(*
SPDX-FileCopyrightText: © 2026 Oleksandr Tiutyk <trofimich@gmail.com>
SPDX-License-Identifier: MIT
License: https://opensource.org/license/mit
*)

(*!
<summary>
Beckhoff EL1512: 2-channel up/down counter terminal (24 V DC).
</summary>
<description>
Represents the default 2Ch. Counter assignment: TxPDOs 0x1A00/0x1A01 and RxPDOs 0x1600/0x1601.
Each channel has 16-bit status/control and a 32-bit counter/preset. Direction is configured through CoE.
Single-channel up/down or gated-counter assignments are outside this model.
When used for I/O, link located fields or their containing buffers to the matching selected PDOs.
The record is not a packed wire buffer; compiler padding is not part of the device specification.
Unlinked/default values do not prove valid I/O. The caller evaluates bus/channel validity before use.
Use one owner task per instance and externally synchronize other access; multi-field snapshots are not atomic.
Copies store data without creating hardware links. Keep borrowed field references valid while consumers are bound.
This passive record performs no validation, synchronization, configuration or protocol advancement.
</description>
*)
TYPE EL1512 :
STRUCT
	Ch1 : COUNTER_CHANNEL;
	Ch2 : COUNTER_CHANNEL;
END_STRUCT
END_TYPE

(* stored: Version 1.1.0.1, ProductVersion 3.1.4026.20
   DUT EL1512: Id {6ce2c619-f95e-46c0-8595-e21364545aac} *)
